// TIA Portal V21 export
// export: Created 2026-10-23T20:43:21.0219718Z, ExportSetting WithDefaults, DisplayName Totally Integrated Automation Portal, DisplayVersion V21 Update 1, DisplayName SINAMICS Startdrive Advanced, DisplayVersion V21 HF2, DisplayName SINAMICS Startdrive G110M, G120, G120C, G120D, G120P, G115D, DisplayVersion V21 HF2, DisplayName SINAMICS Startdrive G130, G150, S120, S150, G200, G220, S200, S210, S220, Innomotics MVD, DisplayVersion V21 HF2, DisplayName STEP 7 Professional, DisplayVersion V21 Update 1, DisplayName STEP 7 Safety, DisplayVersion V21, DisplayName Tech WebApplication, DisplayVersion V21, DisplayName WinCC Basic/Comfort/Advanced, DisplayVersion V21 Update 1, DisplayName WinCC Unified, DisplayVersion V21 Update 1
FUNCTION_BLOCK "FB_AnaGlobalAccess"   // FB14, SCL
TITLE = Analyzer: global access inside an FB
{ S7_Optimized_Access := 'TRUE' }
VERSION : 0.1
// Rule C26g: a global DB and PLC tags are accessed inside the FB
// stored: AutoNumber true, IsIECCheckEnabled false, IsRetainMemResEnabled false, MemoryReserve 100, SetENOAutomatically false, UDAEnableTagReadback false
   VAR_OUTPUT
      Speed : Real;   // Speed setpoint from the global DB
   END_VAR
BEGIN

       #Speed := "DB_Machine".SpeedSetpoint;
       "ConveyorRun" := "StartButton";
END_FUNCTION_BLOCK
